(* IEC 61131-3 sources: llm-plc-st-eval/data/calibracion/claude-sonnet-4-6/B1/few_shot, 3 files *)

(* ---- ejec_1.st ---- *)
```pascal
FUNCTION_BLOCK FB_Motor
VAR_INPUT
    btnMarcha : BOOL; (* Boton de marcha *)
    btnParo   : BOOL; (* Boton de paro *)
    btnEmerg  : BOOL; (* Boton de paro de emergencia *)
END_VAR
VAR_OUTPUT
    motorOn : BOOL; (* Salida del motor *)
END_VAR
VAR
    bloqEmerg : BOOL; (* Bloqueo activo tras paro de emergencia *)
END_VAR

(* Activar bloqueo de emergencia; solo se libera al soltar btnEmerg *)
IF btnEmerg THEN
    bloqEmerg := TRUE;
ELSIF NOT btnEmerg AND NOT btnMarcha THEN
    (* El bloqueo se libera cuando se sueltan emergencia y marcha *)
    bloqEmerg := FALSE;
END_IF;

(* Logica de arranque/paro con autoretencion *)
IF btnParo OR btnEmerg OR bloqEmerg THEN
    (* Paro normal, emergencia o bloqueo activo: apagar motor *)
    motorOn := FALSE;
ELSIF btnMarcha AND NOT bloqEmerg THEN
    (* Arranque: activar motor *)
    motorOn := TRUE;
END_IF;
(* Si ninguna condicion aplica, motorOn conserva su estado (autoretencion) *)

END_FUNCTION_BLOCK
```

(* ---- ejec_2.st ---- *)
```pascal
FUNCTION_BLOCK FB_Motor
VAR_INPUT
    btnMarcha : BOOL; (* Boton de marcha (NA) *)
    btnParo   : BOOL; (* Boton de paro (NC, activo = paro) *)
    btnEmerg  : BOOL; (* Paro de emergencia (NC, activo = emergencia) *)
END_VAR
VAR_OUTPUT
    motorOn : BOOL; (* Contactor / salida del motor *)
END_VAR
VAR
    bloqEmerg : BOOL; (* Bloqueo por emergencia: impide rearranque *)
END_VAR

(* --- Gestion del bloqueo de emergencia --- *)
(* Se activa con btnEmerg y solo se libera cuando btnEmerg vuelve a FALSE *)
(* y el operador no mantiene pulsado btnMarcha (condicion de reset seguro) *)
IF btnEmerg THEN
    bloqEmerg := TRUE;  (* Latch de emergencia *)
ELSIF NOT btnEmerg AND NOT btnMarcha THEN
    bloqEmerg := FALSE; (* Reset del bloqueo solo cuando ambas condiciones son seguras *)
END_IF;

(* --- Logica de arranque / paro con autoretencion --- *)
(* Paro de emergencia o paro normal apagan el motor                        *)
(* El bloqueo impide rearranque tras emergencia aunque btnMarcha este activo *)
IF btnEmerg OR btnParo THEN
    motorOn := FALSE;           (* Paro inmediato por emergencia o paro normal *)
ELSIF btnMarcha AND NOT bloqEmerg THEN
    motorOn := TRUE;            (* Arranque: solo si no hay bloqueo activo *)
END_IF;
(* La autoretencion queda implicita: motorOn mantiene su valor al soltar btnMarcha *)

END_FUNCTION_BLOCK
```

(* ---- ejec_3.st ---- *)
```pascal
FUNCTION_BLOCK FB_Motor
VAR_INPUT
    btnMarcha : BOOL; (* Boton de marcha *)
    btnParo   : BOOL; (* Boton de paro *)
    btnEmerg  : BOOL; (* Boton de paro de emergencia *)
END_VAR
VAR_OUTPUT
    motorOn : BOOL; (* Salida del contactor del motor *)
END_VAR
VAR
    bloqEmerg : BOOL; (* Bloqueo activo tras paro de emergencia *)
END_VAR

(* Activar bloqueo de emergencia; solo se libera al soltar btnEmerg *)
IF btnEmerg THEN
    bloqEmerg := TRUE;
ELSIF NOT btnEmerg AND NOT motorOn THEN
    (* Se libera el bloqueo cuando la emergencia se suelta y el motor esta parado *)
    bloqEmerg := FALSE;
END_IF;

(* Logica de arranque y paro con autoretencion *)
IF btnParo OR btnEmerg OR bloqEmerg THEN
    (* Paro normal, emergencia o bloqueo activo: apagar motor *)
    motorOn := FALSE;
ELSIF btnMarcha AND NOT bloqEmerg THEN
    (* Arranque solo si no hay bloqueo de emergencia *)
    motorOn := TRUE;
END_IF;

END_FUNCTION_BLOCK
```
